{region 'Documentation'}
(*!
<summary>Optional base for a resource Preparation controlled by level-based Enable.</summary>
<description>
Call SUPER^() once per task cycle. Implement Prepare to observe the resource on every call and
perform resource actions only while Enabled.

The base owns the accepted Enable view and status storage, not initialization, a reset
protocol, events or timeout supervision. The Test Case owns the Preparation timeout.

Disabled processing must not issue resource or cleanup commands. Removing Enable does not cancel
an already accepted resource command; the Test Case owns Reset/Abort handling.
</description>
*)
{endregion}
FUNCTION_BLOCK ABSTRACT PreparationBase IMPLEMENTS I_Preparation
VAR_INPUT
    Enable : BOOL; //! Permits resource-changing preparation work; disabled calls may still observe and report the resource.
END_VAR
VAR
    FEnabled : BOOL;
    /// Derived Prepare updates all applicable fields consistently with the Preparation contract.
    FStatus : ST_PreparationStatus;
END_VAR

FEnabled := Enable;
Prepare();

{region 'Documentation'}
(*!
<summary>Enable accepted at the last FB call; not proof of active resource manipulation.</summary>
*)
{endregion}
{attribute 'monitoring' := 'call'}
PROPERTY PUBLIC Enabled : BOOL //! Enable accepted at the last FB call; not proof of active resource manipulation.
GET // PUBLIC
Enabled := FEnabled;
END_GET
END_PROPERTY

{region 'Documentation'}
(*!
<summary>Observes the resource and maintains its Preparation status on every FB call.</summary>
<description>
This abstract hook has no base implementation to call. Use Enabled to gate resource-changing
work; disabled calls must still report current target, readiness and error observations.

On deactivation, stop resource manipulation and return any internal sequence to its executable
base state. Completed reports the current target condition, not a latched success. UpdateStatus may
be used to project consistent flags.
</description>
*)
{endregion}
METHOD PROTECTED ABSTRACT Prepare
END_METHOD

{region 'Documentation'}
(*!
<summary>Snapshot of the status maintained by the concrete Preparation.</summary>
*)
{endregion}
PROPERTY PUBLIC Status : ST_PreparationStatus //! Snapshot of the status maintained by the concrete Preparation.
GET // PUBLIC
Status := FStatus;
END_GET
END_PROPERTY

{region 'Documentation'}
(*!
<summary>Replaces the Preparation snapshot without performing resource work.</summary>
<description>
State is diagnostic context, independent of ExecutionStatus. Running, Completed and Error
follow ExecutionStatus; Ready is suppressed only while Running.

Select E_ExecutionStatus.Idle only when Ready is TRUE and neither work, completion nor error applies; otherwise
select E_ExecutionStatus.NotReady. This method does not validate that choice, latch completion, publish events or
supervise timeouts.
</description>
*)
{endregion}
METHOD PROTECTED UpdateStatus
VAR_INPUT
    State : E_State; //! Concrete Preparation's lifecycle state; independent of the execution-status classification.
    ExecutionStatus : E_ExecutionStatus; //! Execution classification used to derive Running, Completed and Error in the Preparation snapshot.
    Ready : BOOL; //! Resource can be driven to the target state; suppressed while Running. Does not mean target reached.
END_VAR
FStatus.State := State;
FStatus.ExecutionStatus := ExecutionStatus;
FStatus.Running := ExecutionStatus = E_ExecutionStatus.Running;
FStatus.Completed := ExecutionStatus = E_ExecutionStatus.Completed;
FStatus.Error := ExecutionStatus = E_ExecutionStatus.Error;
FStatus.Ready := Ready AND NOT FStatus.Running;
END_METHOD

END_FUNCTION_BLOCK

(* stored: Version 1.1.0.1
   POU PreparationBase: Id {db8d08a6-b7d5-4b1d-aa16-97f6ebd405b3}, SpecialFunc None
   Folder Internal: Id {309f91ec-5692-42b8-9fc2-a08cccea2615}
   Property Enabled: Id {c613fa76-1c4b-4033-8a65-7c9ab2227542}
   Get Get: Id {43451ac6-816b-465e-94f4-17afd4e401c9}
   Method Prepare: Id {2df63df0-2eea-4ccc-89f2-3f965232340e}
   Property Status: Id {d65ca166-f06f-4f93-b34e-47ced876765d}
   Get Get: Id {86be9150-2974-4491-89a6-aa07e276a3ba}
   Method UpdateStatus: Id {def9e459-d79e-4782-8440-002e8559e7bd} *)
